(* IEC 61131-3 sources: virtual-bottling-plant/plc/src/generated/types, 2 files *)

(* ---- Contract_Enums.st ---- *)
(* GENERATED by plc/scripts/gen_plc_io.py from contracts/modbus/plc-io.yaml. Do not edit by hand. *)
(* Enums with fixed contract numbers. matiec enums cannot carry values, so XToInt / IntToX convert at the boundary. *)
TYPE
  E_PackMLState : (PML_UNDEFINED, PML_CLEARING, PML_STOPPED, PML_STARTING, PML_IDLE, PML_SUSPENDED, PML_EXECUTE, PML_STOPPING, PML_ABORTING, PML_ABORTED, PML_HOLDING, PML_HELD, PML_UNHOLDING, PML_SUSPENDING, PML_UNSUSPENDING, PML_RESETTING, PML_COMPLETING, PML_COMPLETE);
  E_PackMLMode : (MODE_NONE, MODE_PRODUCTION, MODE_MAINTENANCE, MODE_MANUAL);
  E_BatchPhase : (PHASE_IDLE, PHASE_FILL, PHASE_MIX, PHASE_TRANSFER, PHASE_DRAIN, PHASE_CIP);
  E_Command : (CMD_NONE, CMD_START, CMD_STOP, CMD_RESET, CMD_ABORT, CMD_CLEAR);
  E_RecipeNak : (NAK_NONE, NAK_IN_EXECUTE, NAK_BRIX_OUT_OF_RANGE, NAK_CONC_RATIO_OUT_OF_RANGE, NAK_FILL_WEIGHT_OUT_OF_RANGE, NAK_LINE_SPEED_OUT_OF_RANGE, NAK_CAP_TORQUE_OUT_OF_RANGE, NAK_UNKNOWN_PRODUCT, NAK_BUSY);
END_TYPE

FUNCTION PackMLStateToInt : INT
  VAR_INPUT
    In : E_PackMLState;
  END_VAR
  CASE In OF
    PML_UNDEFINED: PackMLStateToInt := 0;
    PML_CLEARING: PackMLStateToInt := 1;
    PML_STOPPED: PackMLStateToInt := 2;
    PML_STARTING: PackMLStateToInt := 3;
    PML_IDLE: PackMLStateToInt := 4;
    PML_SUSPENDED: PackMLStateToInt := 5;
    PML_EXECUTE: PackMLStateToInt := 6;
    PML_STOPPING: PackMLStateToInt := 7;
    PML_ABORTING: PackMLStateToInt := 8;
    PML_ABORTED: PackMLStateToInt := 9;
    PML_HOLDING: PackMLStateToInt := 10;
    PML_HELD: PackMLStateToInt := 11;
    PML_UNHOLDING: PackMLStateToInt := 12;
    PML_SUSPENDING: PackMLStateToInt := 13;
    PML_UNSUSPENDING: PackMLStateToInt := 14;
    PML_RESETTING: PackMLStateToInt := 15;
    PML_COMPLETING: PackMLStateToInt := 16;
    PML_COMPLETE: PackMLStateToInt := 17;
  END_CASE;
END_FUNCTION

FUNCTION IntToPackMLState : E_PackMLState
  VAR_INPUT
    In : INT;
  END_VAR
  IntToPackMLState := PML_UNDEFINED;
  CASE In OF
    0: IntToPackMLState := PML_UNDEFINED;
    1: IntToPackMLState := PML_CLEARING;
    2: IntToPackMLState := PML_STOPPED;
    3: IntToPackMLState := PML_STARTING;
    4: IntToPackMLState := PML_IDLE;
    5: IntToPackMLState := PML_SUSPENDED;
    6: IntToPackMLState := PML_EXECUTE;
    7: IntToPackMLState := PML_STOPPING;
    8: IntToPackMLState := PML_ABORTING;
    9: IntToPackMLState := PML_ABORTED;
    10: IntToPackMLState := PML_HOLDING;
    11: IntToPackMLState := PML_HELD;
    12: IntToPackMLState := PML_UNHOLDING;
    13: IntToPackMLState := PML_SUSPENDING;
    14: IntToPackMLState := PML_UNSUSPENDING;
    15: IntToPackMLState := PML_RESETTING;
    16: IntToPackMLState := PML_COMPLETING;
    17: IntToPackMLState := PML_COMPLETE;
  END_CASE;
END_FUNCTION

FUNCTION PackMLModeToInt : INT
  VAR_INPUT
    In : E_PackMLMode;
  END_VAR
  CASE In OF
    MODE_NONE: PackMLModeToInt := 0;
    MODE_PRODUCTION: PackMLModeToInt := 1;
    MODE_MAINTENANCE: PackMLModeToInt := 2;
    MODE_MANUAL: PackMLModeToInt := 3;
  END_CASE;
END_FUNCTION

FUNCTION IntToPackMLMode : E_PackMLMode
  VAR_INPUT
    In : INT;
  END_VAR
  IntToPackMLMode := MODE_NONE;
  CASE In OF
    0: IntToPackMLMode := MODE_NONE;
    1: IntToPackMLMode := MODE_PRODUCTION;
    2: IntToPackMLMode := MODE_MAINTENANCE;
    3: IntToPackMLMode := MODE_MANUAL;
  END_CASE;
END_FUNCTION

FUNCTION BatchPhaseToInt : INT
  VAR_INPUT
    In : E_BatchPhase;
  END_VAR
  CASE In OF
    PHASE_IDLE: BatchPhaseToInt := 0;
    PHASE_FILL: BatchPhaseToInt := 1;
    PHASE_MIX: BatchPhaseToInt := 2;
    PHASE_TRANSFER: BatchPhaseToInt := 3;
    PHASE_DRAIN: BatchPhaseToInt := 4;
    PHASE_CIP: BatchPhaseToInt := 5;
  END_CASE;
END_FUNCTION

FUNCTION IntToBatchPhase : E_BatchPhase
  VAR_INPUT
    In : INT;
  END_VAR
  IntToBatchPhase := PHASE_IDLE;
  CASE In OF
    0: IntToBatchPhase := PHASE_IDLE;
    1: IntToBatchPhase := PHASE_FILL;
    2: IntToBatchPhase := PHASE_MIX;
    3: IntToBatchPhase := PHASE_TRANSFER;
    4: IntToBatchPhase := PHASE_DRAIN;
    5: IntToBatchPhase := PHASE_CIP;
  END_CASE;
END_FUNCTION

FUNCTION CommandToInt : INT
  VAR_INPUT
    In : E_Command;
  END_VAR
  CASE In OF
    CMD_NONE: CommandToInt := 0;
    CMD_START: CommandToInt := 1;
    CMD_STOP: CommandToInt := 2;
    CMD_RESET: CommandToInt := 3;
    CMD_ABORT: CommandToInt := 4;
    CMD_CLEAR: CommandToInt := 5;
  END_CASE;
END_FUNCTION

FUNCTION IntToCommand : E_Command
  VAR_INPUT
    In : INT;
  END_VAR
  IntToCommand := CMD_NONE;
  CASE In OF
    0: IntToCommand := CMD_NONE;
    1: IntToCommand := CMD_START;
    2: IntToCommand := CMD_STOP;
    3: IntToCommand := CMD_RESET;
    4: IntToCommand := CMD_ABORT;
    5: IntToCommand := CMD_CLEAR;
  END_CASE;
END_FUNCTION

FUNCTION RecipeNakToInt : INT
  VAR_INPUT
    In : E_RecipeNak;
  END_VAR
  CASE In OF
    NAK_NONE: RecipeNakToInt := 0;
    NAK_IN_EXECUTE: RecipeNakToInt := 1;
    NAK_BRIX_OUT_OF_RANGE: RecipeNakToInt := 2;
    NAK_CONC_RATIO_OUT_OF_RANGE: RecipeNakToInt := 3;
    NAK_FILL_WEIGHT_OUT_OF_RANGE: RecipeNakToInt := 4;
    NAK_LINE_SPEED_OUT_OF_RANGE: RecipeNakToInt := 5;
    NAK_CAP_TORQUE_OUT_OF_RANGE: RecipeNakToInt := 6;
    NAK_UNKNOWN_PRODUCT: RecipeNakToInt := 7;
    NAK_BUSY: RecipeNakToInt := 8;
  END_CASE;
END_FUNCTION

FUNCTION IntToRecipeNak : E_RecipeNak
  VAR_INPUT
    In : INT;
  END_VAR
  IntToRecipeNak := NAK_NONE;
  CASE In OF
    0: IntToRecipeNak := NAK_NONE;
    1: IntToRecipeNak := NAK_IN_EXECUTE;
    2: IntToRecipeNak := NAK_BRIX_OUT_OF_RANGE;
    3: IntToRecipeNak := NAK_CONC_RATIO_OUT_OF_RANGE;
    4: IntToRecipeNak := NAK_FILL_WEIGHT_OUT_OF_RANGE;
    5: IntToRecipeNak := NAK_LINE_SPEED_OUT_OF_RANGE;
    6: IntToRecipeNak := NAK_CAP_TORQUE_OUT_OF_RANGE;
    7: IntToRecipeNak := NAK_UNKNOWN_PRODUCT;
    8: IntToRecipeNak := NAK_BUSY;
  END_CASE;
END_FUNCTION

(* ---- Contract_Structs.st ---- *)
(* GENERATED by plc/scripts/gen_plc_io.py from contracts/modbus/sim-io.yaml + plc-io.yaml. Do not edit by hand. *)
(* Process image (sim I/O in engineering units) and bridge structs. *)
TYPE
  ST_SimInputs : STRUCT
    LT101_Level : REAL;
    AT101_Brix : REAL;
    FT101_WaterFlow : REAL;
    FT102_ConcFlow : REAL;
    FT103_SugarFlow : REAL;
    ST101_AgitatorRpm : REAL;
    T101_ConcLotNo : UDINT;
    T101_Heartbeat : UINT;
    LSL101_Empty : BOOL;
    M101_Running : BOOL;
    T101_CipDone : BOOL;
    TT201_InTemp : REAL;
    TT202_OutTemp : REAL;
    FT201_Flow : REAL;
    PT201_SteamPressure : REAL;
    P201_Heartbeat : UINT;
    ZS203_DivertOpen : BOOL;
    LT301_Level : REAL;
    T301_Heartbeat : UINT;
    LSL301_Low : BOOL;
    F401_Speed : REAL;
    F401_Count : UDINT;
    F401_Heartbeat : UINT;
    F401_Running : BOOL;
    F401_NozzleLeak : BOOL;
    C501_Speed : REAL;
    C501_Count : UDINT;
    C501_Torque : REAL;
    LT502_CapHopper : REAL;
    C501_Heartbeat : UINT;
    C501_Running : BOOL;
    C501_Jam : BOOL;
    C501_Breakdown : BOOL;
    LSL502_CapsEmpty : BOOL;
    L601_Speed : REAL;
    L601_Count : UDINT;
    L601_RollRemaining : REAL;
    L601_Heartbeat : UINT;
    L601_Running : BOOL;
    L601_RollEmpty : BOOL;
    L601_LabelError : BOOL;
    L601_Breakdown : BOOL;
    Q701_Speed : REAL;
    Q701_Count : UDINT;
    Q701_RejectCount : UDINT;
    WT701_LastWeight : REAL;
    Q701_Heartbeat : UINT;
    Q701_N01_Seq : UINT;
    Q701_N01_Mean : REAL;
    Q701_N01_Range : REAL;
    Q701_N02_Seq : UINT;
    Q701_N02_Mean : REAL;
    Q701_N02_Range : REAL;
    Q701_N03_Seq : UINT;
    Q701_N03_Mean : REAL;
    Q701_N03_Range : REAL;
    Q701_N04_Seq : UINT;
    Q701_N04_Mean : REAL;
    Q701_N04_Range : REAL;
    Q701_N05_Seq : UINT;
    Q701_N05_Mean : REAL;
    Q701_N05_Range : REAL;
    Q701_N06_Seq : UINT;
    Q701_N06_Mean : REAL;
    Q701_N06_Range : REAL;
    Q701_N07_Seq : UINT;
    Q701_N07_Mean : REAL;
    Q701_N07_Range : REAL;
    Q701_N08_Seq : UINT;
    Q701_N08_Mean : REAL;
    Q701_N08_Range : REAL;
    Q701_N09_Seq : UINT;
    Q701_N09_Mean : REAL;
    Q701_N09_Range : REAL;
    Q701_N10_Seq : UINT;
    Q701_N10_Mean : REAL;
    Q701_N10_Range : REAL;
    Q701_N11_Seq : UINT;
    Q701_N11_Mean : REAL;
    Q701_N11_Range : REAL;
    Q701_N12_Seq : UINT;
    Q701_N12_Mean : REAL;
    Q701_N12_Range : REAL;
    Q701_Running : BOOL;
    K801_Speed : REAL;
    K801_CaseCount : UDINT;
    K801_Heartbeat : UINT;
    K801_Running : BOOL;
    K801_Jam : BOOL;
    K801_Breakdown : BOOL;
    SIM_TimeMs : UDINT;
    CV1_Fill : REAL;
    CV2_Fill : REAL;
    CV3_Fill : REAL;
    CV4_Fill : REAL;
    LINE_Heartbeat : UINT;
    CV1_Full : BOOL;
    CV2_Full : BOOL;
    CV3_Full : BOOL;
    CV4_Full : BOOL;
    PB_Start : BOOL;
    PB_Stop : BOOL;
    PB_Reset : BOOL;
  END_STRUCT;
  ST_SimOutputs : STRUCT
    XV101_Water : BOOL;
    XV102_Conc : BOOL;
    XV103_Sugar : BOOL;
    M101_Agitator : BOOL;
    P101_TransferPump : BOOL;
    XV109_Drain : BOOL;
    T101_CipRun : BOOL;
    T101_ConcSelect : REAL;
    XV203_Divert : BOOL;
    TCV201_SteamValve : REAL;
    XV309_Drain : BOOL;
    F401_Run : BOOL;
    F401_SpeedSP : REAL;
    F401_FillTargetG : REAL;
    C501_Run : BOOL;
    C501_SpeedSP : REAL;
    L601_Run : BOOL;
    L601_SpeedSP : REAL;
    Q701_Run : BOOL;
    Q701_SpeedSP : REAL;
    Q701_RejectLimitG : REAL;
    K801_Run : BOOL;
    K801_SpeedSP : REAL;
  END_STRUCT;
  ST_T101Status : STRUCT
    Phase : E_BatchPhase;
    BatchNo : INT;
    ProductCode : INT;
    BatchBrix : REAL;
    BrixOk : BOOL;
    BatchActive : BOOL;
  END_STRUCT;
  ST_P201Status : STRUCT
    TempSP : REAL;
    DivertCount : INT;
    ForwardFlowOk : BOOL;
  END_STRUCT;
  ST_T301Status : STRUCT
    FillerPermissive : BOOL;
  END_STRUCT;
  ST_PackagingStatus : STRUCT
    State : E_PackMLState;
    Mode : E_PackMLMode;
    StopReason : INT;
    Blocked : BOOL;
    Starved : BOOL;
  END_STRUCT;
  ST_LINEStatus : STRUCT
    State : E_PackMLState;
    RecipeId : INT;
    RecipeVersion : INT;
    ProductCode : INT;
    PlcHeartbeat : INT;
  END_STRUCT;
  ST_Status : STRUCT
    T101 : ST_T101Status;
    P201 : ST_P201Status;
    T301 : ST_T301Status;
    F401 : ST_PackagingStatus;
    C501 : ST_PackagingStatus;
    L601 : ST_PackagingStatus;
    Q701 : ST_PackagingStatus;
    K801 : ST_PackagingStatus;
    LINE : ST_LINEStatus;
  END_STRUCT;
  ST_CommsStatus : STRUCT
    T101 : BOOL;
    P201 : BOOL;
    T301 : BOOL;
    F401 : BOOL;
    C501 : BOOL;
    L601 : BOOL;
    Q701 : BOOL;
    K801 : BOOL;
    LINE : BOOL;
  END_STRUCT;
  ST_AlarmSummary : STRUCT
    T101_Word : INT;
    P201_Word : INT;
    T301_Word : INT;
    F401_Word : INT;
    C501_Word : INT;
    L601_Word : INT;
    Q701_Word : INT;
    K801_Word : INT;
    LINE_Word : INT;
    T101_ActiveId : INT;
    P201_ActiveId : INT;
    T301_ActiveId : INT;
    F401_ActiveId : INT;
    C501_ActiveId : INT;
    L601_ActiveId : INT;
    Q701_ActiveId : INT;
    K801_ActiveId : INT;
    LINE_ActiveId : INT;
    ActiveCount : INT;
    FirstOutId : INT;
    W1 : UINT;
    W2 : UINT;
    W3 : UINT;
    W4 : UINT;
    W5 : UINT;
    W6 : UINT;
    W7 : UINT;
    W8 : UINT;
    W9 : UINT;
    W10 : UINT;
    W11 : UINT;
    W12 : UINT;
    W13 : UINT;
    W14 : UINT;
    W15 : UINT;
    W16 : UINT;
    W17 : UINT;
    W18 : UINT;
    W19 : UINT;
    W20 : UINT;
    W21 : UINT;
    W22 : UINT;
  END_STRUCT;
  ST_Counters : STRUCT
    Q701_GoodCount : UDINT;
  END_STRUCT;
  ST_Commands : STRUCT
    F401_Cmd : E_Command;
    C501_Cmd : E_Command;
    L601_Cmd : E_Command;
    Q701_Cmd : E_Command;
    K801_Cmd : E_Command;
    LINE_Cmd : E_Command;
    F401_StopReason : INT;
    C501_StopReason : INT;
    L601_StopReason : INT;
    Q701_StopReason : INT;
    K801_StopReason : INT;
    AlarmAck : INT;
    P201_TempSP : REAL;
  END_STRUCT;
  ST_RecipeRequest : STRUCT
    Recipe_Req : BOOL;
    RecipeId : INT;
    RecipeVersion : INT;
    ProductCode : INT;
    BrixTarget : REAL;
    BrixTol : REAL;
    ConcRatio : REAL;
    FillTargetG : REAL;
    LineSpeed : INT;
    CapTorque : REAL;
  END_STRUCT;
  ST_RecipeResponse : STRUCT
    Recipe_Ack : BOOL;
    Recipe_Nak : E_RecipeNak;
  END_STRUCT;
END_TYPE
